Staubli VAL3: initList.pgx

public program initList(utList& x_utList[], string x_sPage, string x_sId)
begin
  x_utList.Common.sPage=x_sPage
  x_utList.Common.sID=x_sId
  userPageBind(x_utList.Common.sPage,x_utList.Common.sID,"options",x_utList.Common.sItem,size(x_utList.Common.sItem),"r")
  userPageBind(x_utList.Common.sPage,x_utList.Common.sID,"value",x_utList.Common.sValue,1,"rw")
end
